{attribute 'pack_mode' := '1'}
TYPE ST_PcsPublishData :
STRUCT
	Header		:	ST_MqttHeader;
	Devices		:	ARRAY[0..GVL_PARAM.PCS_COUNT-1] OF ST_PcsPublish_V1;
END_STRUCT
END_TYPE

(* stored: Version 1.1.0.1, ProductVersion 3.1.4024.15
   DUT ST_PcsPublishData: Id {ae5bcb89-b667-4961-8d48-231ab80d5344} *)
